(* PLC project zarechnaya.project, CODESYS CODESYS V3.5 SP17 Patch 3 *)
(* stored: creationDateTime 2026-10-20T05:42:22.2568826, modificationDateTime 1601-01-01T03:00:00 *)

(* FB_PiCfc — ПИ-регулятор расхода промывочной воды (CFC, обратная связь). Поведение (модель scenarios/reference/model_FB_PiCfc.py), шаги executionOrderId: 1. e := rSp − rPv; 2. p := rKp · e; 3. k := rKi · e; 4. i := k + i (вход In2 блока ADD — его собственный выход: значение прошлого цикла, начально 0; C2S7-GFX-CFCFB); 5. u := p + i; 6. o := LIMIT(rMin, u, rMax); 7. rOut := o. Все операции — REAL (float32). *)
FUNCTION_BLOCK FB_PiCfc
  VAR_INPUT
    rSp : REAL;
    rPv : REAL;
    rKp : REAL;
    rKi : REAL;
    rMin : REAL;
    rMax : REAL;
  END_VAR
  VAR_OUTPUT
    rOut : REAL;
  END_VAR
  VAR  (* added by the conversion: wires and edge detectors of the diagram *)
    _SUB11_OUT : REAL;
    _ADD17_OUT : ANY;
  END_VAR

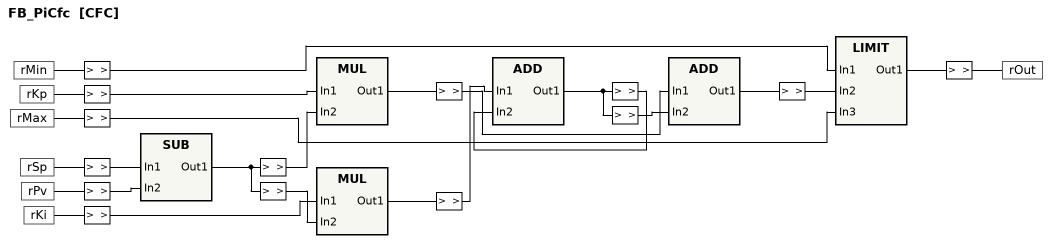
(* CFC diagram, written out as Structured Text *)
_SUB11_OUT := rSp - rPv;
_ADD17_OUT := rKi * _SUB11_OUT + _ADD17_OUT;
rOut := LIMIT(rMin, rKp * _SUB11_OUT + _ADD17_OUT, rMax);
END_FUNCTION_BLOCK
